INTERFACE I_IoBit EXTENDS I_IoBase

PROPERTY ftrig : BOOL
GET
END_GET
SET
END_SET
END_PROPERTY

PROPERTY Q : BOOL
GET
END_GET
SET
END_SET
END_PROPERTY

PROPERTY rtrig : BOOL
GET
END_GET
SET
END_SET
END_PROPERTY

END_INTERFACE

(* stored: Version 1.1.0.1
   Itf I_IoBit: Id {4c8a557e-4677-4e4f-a074-934e8ef598b1}
   Property ftrig: Id {36b1dff4-b3a6-455b-b902-afb68be29cdd}
   Get Get: Id {e2da75fc-c981-4453-b59b-593dcaa3c7a9}
   Set Set: Id {89f6fb45-35d5-44c4-b642-3de7a7505330}
   Property Q: Id {d840fc8f-f573-47e4-9e5f-3d3ad7a79148}
   Get Get: Id {4d4b5465-6152-46ae-a729-07dc9aa06957}
   Set Set: Id {e6eeaf8d-ae0c-483b-a3c5-db6fa4ec7717}
   Property rtrig: Id {cc3d6f26-b3e3-494e-a9ae-0100b97b793a}
   Get Get: Id {c23d3a32-ed0d-4544-b194-34f61f6b2fb4}
   Set Set: Id {3aa53ac3-3cd3-4ea3-91e9-16d3fd112db7} *)
